(* IEC 61131-3 sources: volt/packages/volt-lsp-iec/test-corpus/pro2193/Device/Plc Logic/Application/99 Library/Functions/PositionReached, 2 files *)

(* ---- PositionReached.pou ---- *)
// Check if two positions match (within 1 mm).
FUNCTION PositionReached : BOOL
VAR_INPUT
	rActPos		: REAL;
	rSetPos		: REAL;
END_VAR

%LANGUAGE ST
PositionReached			:= PositionReachedValue(rActPos, rSetPos, 1);

END_FUNCTION

(* ---- PositionReachedValue.pou ---- *)
// Check if two positions match (within rValue mm).
FUNCTION PositionReachedValue : BOOL
VAR_INPUT
	rActPos		: REAL;
	rSetPos		: REAL;
	rValue		: REAL;
END_VAR

%LANGUAGE ST
PositionReachedValue	:= ABS(rActPos - rSetPos) <= rValue;

END_FUNCTION
